Staubli VAL3: getDigIO.pgx

public program getDigIO(dio x_dIO, bool& x_bValue, bool& x_bError)
  local string l_sDesc
  local string l_sPath
begin
  if ioStatus(x_dIO,l_sDesc,l_sPath)>=0
    x_bError=false
    x_bValue=(x_dIO==true)
  else
    x_bError=true
  endIf
end
